(* IEC 61131-3 sources: CNC-Cell-Simulator/source/plc (part 2) *)

PROGRAM CellMain
  VAR_EXTERNAL
    R1_state : INT;
    R1_fault : INT;
    CONV_state : INT;
    CONV_fault : INT;
    R2_state : INT;
    R2_fault : INT;
    SUP_state : INT;
    SAF_state : INT;
    R1_JobNo : INT;
    R1_Start : BOOL;
    R1_Done : BOOL;
    R1_CP_1_Trig : BOOL;
    R1_CP_1_Done : BOOL;
    R1_CP_1_Valid : BOOL;
    R1_CP_1_Cam : BOOL;
    R1_CP_1_Also : BOOL;
    R1_CP_2_Trig : BOOL;
    R1_CP_2_Done : BOOL;
    R1_CP_2_Valid : BOOL;
    R1_CP_2_Cam : BOOL;
    CONV_CP_2_Trig : BOOL;
    CONV_CP_2_Done : BOOL;
    CONV_CP_2_Valid : BOOL;
    CONV_CP_2_Cam : BOOL;
    CONV_CP_3_Trig : BOOL;
    CONV_CP_3_Done : BOOL;
    CONV_CP_3_Valid : BOOL;
    CONV_CP_3_Cam : BOOL;
    R2_JobNo : INT;
    R2_Start : BOOL;
    R2_Done : BOOL;
    R2_CP_4_Trig : BOOL;
    R2_CP_4_Done : BOOL;
    R2_CP_4_Valid : BOOL;
    R2_CP_4_Cam : BOOL;
    R2_CP_5_Trig : BOOL;
    R2_CP_5_Done : BOOL;
    R2_CP_5_Valid : BOOL;
    R2_CP_5_Cam : BOOL;
    R2_CP_3_Trig : BOOL;
    R2_CP_3_Done : BOOL;
    R2_CP_3_Valid : BOOL;
    R2_CP_3_Cam : BOOL;
    HMI_auto : BOOL;
    R1_home : BOOL;
    CNC_ready : BOOL;
    ZS_32_in : BOOL;
    ZS_32 : BOOL;
    SC_01_prot : BOOL;
    GR_21A_in : BOOL;
    GR_21A : BOOL;
    CNC_done : BOOL;
    CNC_empty : BOOL;
    ZS_33_in : BOOL;
    ZS_33 : BOOL;
    ZS_31_in : BOOL;
    ZS_31 : BOOL;
    PS_36_in : BOOL;
    PS_36 : BOOL;
    GR_21B_in : BOOL;
    GR_21B : BOOL;
    ZS_34_in : BOOL;
    ZS_34 : BOOL;
    ZS_35_in : BOOL;
    ZS_35 : BOOL;
    R1_clearCnc : BOOL;
    CNC_run : BOOL;
    ENC_43_in : BOOL;
    ENC_43 : BOOL;
    R1_clearConv : BOOL;
    HMI_loaded : BOOL;
    R2_clearConv : BOOL;
    PE_42_in : BOOL;
    PE_42 : BOOL;
    ROI_C : BOOL;
    R2_home : BOOL;
    GAUGE_zeroed : BOOL;
    GAUGE_due : BOOL;
    GAUGE_due_restart : BOOL;
    GR_51_in : BOOL;
    GR_51 : BOOL;
    R2_clearGauge : BOOL;
    GAUGE_valid : BOOL;
    GAUGE_ok : BOOL;
    SC_02_prot : BOOL;
    CAM_2_slot : BOOL;
    outCount : INT;
    PE_65_in : BOOL;
    PE_65 : BOOL;
    ESTOP : BOOL;
    R1_safeStop : BOOL;
    R2_safeStop : BOOL;
    SC_01_warn : BOOL;
    SC_02_warn : BOOL;
    GAUGE_warn : BOOL;
    PX_11_in : BOOL;
    PX_11 : BOOL;
    PE_41_in : BOOL;
    PE_41 : BOOL;
    PX_52_in : BOOL;
    PX_52 : BOOL;
    PX_64_in : BOOL;
    PX_64 : BOOL;
    HMI_clear : BOOL;
    E_HMI_clear : BOOL;
    HMI_verify : BOOL;
    L_HMI_verify : BOOL;
    VERIFY_pass : BOOL;
    L_VERIFY_pass : BOOL;
    HMI_reset : BOOL;
    L_HMI_reset : BOOL;
    VERIFY_fail : BOOL;
    L_VERIFY_fail : BOOL;
    HMI_safety : BOOL;
    L_HMI_safety : BOOL;
    HMI_release : BOOL;
    L_HMI_release : BOOL;
    HMI_tool : BOOL;
    L_HMI_tool : BOOL;
    HB : BOOL;
    partPlaced : BOOL;
    pickAllowed : BOOL;
    partPicked : BOOL;
    consecNok : INT;
    QH : BOOL;
    toolCount : INT;
    mismatches : INT;
    CAM_FAULT : BOOL;
    COMM_LOST : BOOL;
    mmPending : INT;
    mmClear : BOOL;
    BELT_motor : BOOL;
    LT_53 : BOOL;
    LT_01_red : BOOL;
    LT_01_amber : BOOL;
    LT_01_green : BOOL;
    V_partPlaced : BOOL;
    V_pickAllowed : BOOL;
    V_partPicked : BOOL;
    V_consecNok : INT;
    V_QH : BOOL;
    V_toolCount : INT;
    V_mismatches : INT;
    V_CAM_FAULT : BOOL;
    TR_N : INT;
    TR_00 : INT;
    TR_01 : INT;
    TR_02 : INT;
    TR_03 : INT;
    TR_04 : INT;
    TR_05 : INT;
    TR_06 : INT;
    TR_07 : INT;
    TR_08 : INT;
    TR_09 : INT;
    TR_10 : INT;
    TR_11 : INT;
    TR_12 : INT;
    TR_13 : INT;
    TR_14 : INT;
    TR_15 : INT;
    TR_16 : INT;
    TR_17 : INT;
    TR_18 : INT;
    TR_19 : INT;
    TR_20 : INT;
    TR_21 : INT;
    TR_22 : INT;
    TR_23 : INT;
    TR_24 : INT;
    TR_25 : INT;
    TR_26 : INT;
    TR_27 : INT;
    TR_28 : INT;
    TR_29 : INT;
    TR_30 : INT;
    TR_31 : INT;
  END_VAR
  VAR
    fbR1S2 : FB_R1S2;
    fbCONV : FB_CONV;
    fbR2S2 : FB_R2S2;
    fbSUP : FB_SUP;
    fbSAF : FB_SAF;
    hbT : TON;
    hbLast : BOOL;
    n : INT;
    oldest : INT;
    best : TIME;
    db_ZS_32 : TON;
    db_GR_21A : TON;
    db_ZS_33 : TON;
    db_ZS_31 : TON;
    db_PS_36 : TON;
    db_GR_21B : TON;
    db_ZS_34 : TON;
    db_ZS_35 : TON;
    db_ENC_43 : TON;
    db_PE_42 : TON;
    db_GR_51 : TON;
    db_PX_11 : TON;
    db_PE_41 : TON;
    db_PX_52 : TON;
    db_PX_64 : TON;
    rt_PE_65 : R_TRIG;
    rt_HMI_clear : R_TRIG;
    rt_HMI_verify : R_TRIG;
    rt_VERIFY_pass : R_TRIG;
    rt_HMI_reset : R_TRIG;
    rt_VERIFY_fail : R_TRIG;
    rt_HMI_safety : R_TRIG;
    rt_HMI_release : R_TRIG;
    rt_HMI_tool : R_TRIG;
    mmOn1 : BOOL;
    mmT1 : TON;
    mmOn2 : BOOL;
    mmT2 : TON;
    mmOn3 : BOOL;
    mmT3 : TON;
    tm_GAUGE_due : TON;
    trBuf : ARRAY[0..31] OF INT;
    trI : INT;
    trL_R1 : INT;
    trL_CONV : INT;
    trL_R2 : INT;
    trL_SUP : INT;
    trL_SAF : INT;
  END_VAR
  (* 1. inputs: heartbeat, debounce, latches, mismatch window, PLC timers *)
  hbT(IN := HB = hbLast, PT := T#500ms); hbLast := HB; COMM_LOST := hbT.Q;
  db_ZS_32(IN := ZS_32_in <> ZS_32, PT := T#50ms); IF db_ZS_32.Q THEN ZS_32 := ZS_32_in; END_IF;
  db_GR_21A(IN := GR_21A_in <> GR_21A, PT := T#50ms); IF db_GR_21A.Q THEN GR_21A := GR_21A_in; END_IF;
  db_ZS_33(IN := ZS_33_in <> ZS_33, PT := T#50ms); IF db_ZS_33.Q THEN ZS_33 := ZS_33_in; END_IF;
  db_ZS_31(IN := ZS_31_in <> ZS_31, PT := T#50ms); IF db_ZS_31.Q THEN ZS_31 := ZS_31_in; END_IF;
  db_PS_36(IN := PS_36_in <> PS_36, PT := T#50ms); IF db_PS_36.Q THEN PS_36 := PS_36_in; END_IF;
  db_GR_21B(IN := GR_21B_in <> GR_21B, PT := T#50ms); IF db_GR_21B.Q THEN GR_21B := GR_21B_in; END_IF;
  db_ZS_34(IN := ZS_34_in <> ZS_34, PT := T#50ms); IF db_ZS_34.Q THEN ZS_34 := ZS_34_in; END_IF;
  db_ZS_35(IN := ZS_35_in <> ZS_35, PT := T#50ms); IF db_ZS_35.Q THEN ZS_35 := ZS_35_in; END_IF;
  db_ENC_43(IN := ENC_43_in <> ENC_43, PT := T#50ms); IF db_ENC_43.Q THEN ENC_43 := ENC_43_in; END_IF;
  db_PE_42(IN := PE_42_in <> PE_42, PT := T#50ms); IF db_PE_42.Q THEN PE_42 := PE_42_in; END_IF;
  db_GR_51(IN := GR_51_in <> GR_51, PT := T#50ms); IF db_GR_51.Q THEN GR_51 := GR_51_in; END_IF;
  db_PX_11(IN := PX_11_in <> PX_11, PT := T#50ms); IF db_PX_11.Q THEN PX_11 := PX_11_in; END_IF;
  db_PE_41(IN := PE_41_in <> PE_41, PT := T#50ms); IF db_PE_41.Q THEN PE_41 := PE_41_in; END_IF;
  db_PX_52(IN := PX_52_in <> PX_52, PT := T#50ms); IF db_PX_52.Q THEN PX_52 := PX_52_in; END_IF;
  db_PX_64(IN := PX_64_in <> PX_64, PT := T#50ms); IF db_PX_64.Q THEN PX_64 := PX_64_in; END_IF;
  rt_PE_65(CLK := PE_65_in); IF rt_PE_65.Q THEN PE_65 := TRUE; END_IF;
  rt_HMI_clear(CLK := HMI_clear); E_HMI_clear := rt_HMI_clear.Q;
  rt_HMI_verify(CLK := HMI_verify); IF rt_HMI_verify.Q THEN L_HMI_verify := TRUE; END_IF;
  rt_VERIFY_pass(CLK := VERIFY_pass); IF rt_VERIFY_pass.Q THEN L_VERIFY_pass := TRUE; END_IF;
  rt_HMI_reset(CLK := HMI_reset); IF rt_HMI_reset.Q THEN L_HMI_reset := TRUE; END_IF;
  rt_VERIFY_fail(CLK := VERIFY_fail); IF rt_VERIFY_fail.Q THEN L_VERIFY_fail := TRUE; END_IF;
  rt_HMI_safety(CLK := HMI_safety); IF rt_HMI_safety.Q THEN L_HMI_safety := TRUE; END_IF;
  rt_HMI_release(CLK := HMI_release); IF rt_HMI_release.Q THEN L_HMI_release := TRUE; END_IF;
  rt_HMI_tool(CLK := HMI_tool); IF rt_HMI_tool.Q THEN L_HMI_tool := TRUE; END_IF;
  IF mmClear THEN mmOn1 := FALSE; mmOn2 := FALSE; mmOn3 := FALSE; mmClear := FALSE; END_IF;
  WHILE mmPending > 0 DO (* a new mismatch event: a free place, or the oldest one is replaced *)
    oldest := 0; best := T#0ms;
    IF oldest >= 0 AND NOT mmOn1 THEN oldest := -1; ELSIF oldest >= 0 AND mmT1.ET >= best THEN best := mmT1.ET; oldest := 1; END_IF;
    IF oldest >= 0 AND NOT mmOn2 THEN oldest := -2; ELSIF oldest >= 0 AND mmT2.ET >= best THEN best := mmT2.ET; oldest := 2; END_IF;
    IF oldest >= 0 AND NOT mmOn3 THEN oldest := -3; ELSIF oldest >= 0 AND mmT3.ET >= best THEN best := mmT3.ET; oldest := 3; END_IF;
    IF oldest < 0 THEN oldest := -oldest; END_IF;
    IF oldest = 1 THEN mmOn1 := TRUE; mmT1(IN := FALSE); END_IF;
    IF oldest = 2 THEN mmOn2 := TRUE; mmT2(IN := FALSE); END_IF;
    IF oldest = 3 THEN mmOn3 := TRUE; mmT3(IN := FALSE); END_IF;
    mmPending := mmPending - 1;
  END_WHILE;
  n := 0;
  mmT1(IN := mmOn1, PT := T#600000ms); IF mmT1.Q THEN mmOn1 := FALSE; mmT1(IN := FALSE); END_IF; IF mmOn1 THEN n := n + 1; END_IF;
  mmT2(IN := mmOn2, PT := T#600000ms); IF mmT2.Q THEN mmOn2 := FALSE; mmT2(IN := FALSE); END_IF; IF mmOn2 THEN n := n + 1; END_IF;
  mmT3(IN := mmOn3, PT := T#600000ms); IF mmT3.Q THEN mmOn3 := FALSE; mmT3(IN := FALSE); END_IF; IF mmOn3 THEN n := n + 1; END_IF;
  mismatches := n;
  IF GAUGE_due_restart THEN tm_GAUGE_due(IN := FALSE); GAUGE_due_restart := FALSE; END_IF;
  tm_GAUGE_due(IN := GAUGE_zeroed, PT := T#14400000ms); GAUGE_due := tm_GAUGE_due.Q;

  (* 2. machines in a fixed order; the urgent supervisor first and after every other machine *)
  fbSUP(); IF SUP_state <> trL_SUP THEN trL_SUP := SUP_state; trBuf[trI MOD 32] := 400 + SUP_state; trI := trI + 1; IF trI >= 32000 THEN trI := 0; END_IF; END_IF;
  fbSAF(); IF SAF_state <> trL_SAF THEN trL_SAF := SAF_state; trBuf[trI MOD 32] := 500 + SAF_state; trI := trI + 1; IF trI >= 32000 THEN trI := 0; END_IF; END_IF;
  fbR1S2(); IF R1_state <> trL_R1 THEN trL_R1 := R1_state; trBuf[trI MOD 32] := 100 + R1_state; trI := trI + 1; IF trI >= 32000 THEN trI := 0; END_IF; END_IF;
  fbSUP(); IF SUP_state <> trL_SUP THEN trL_SUP := SUP_state; trBuf[trI MOD 32] := 400 + SUP_state; trI := trI + 1; IF trI >= 32000 THEN trI := 0; END_IF; END_IF;
  fbSAF(); IF SAF_state <> trL_SAF THEN trL_SAF := SAF_state; trBuf[trI MOD 32] := 500 + SAF_state; trI := trI + 1; IF trI >= 32000 THEN trI := 0; END_IF; END_IF;
  fbCONV(); IF CONV_state <> trL_CONV THEN trL_CONV := CONV_state; trBuf[trI MOD 32] := 200 + CONV_state; trI := trI + 1; IF trI >= 32000 THEN trI := 0; END_IF; END_IF;
  fbSUP(); IF SUP_state <> trL_SUP THEN trL_SUP := SUP_state; trBuf[trI MOD 32] := 400 + SUP_state; trI := trI + 1; IF trI >= 32000 THEN trI := 0; END_IF; END_IF;
  fbSAF(); IF SAF_state <> trL_SAF THEN trL_SAF := SAF_state; trBuf[trI MOD 32] := 500 + SAF_state; trI := trI + 1; IF trI >= 32000 THEN trI := 0; END_IF; END_IF;
  fbR2S2(); IF R2_state <> trL_R2 THEN trL_R2 := R2_state; trBuf[trI MOD 32] := 300 + R2_state; trI := trI + 1; IF trI >= 32000 THEN trI := 0; END_IF; END_IF;
  IF (L_HMI_release AND QH) THEN QH := FALSE; consecNok := 0; L_HMI_release := FALSE; END_IF; (* rung: tool and offsets checked -> quality hold released *)
  IF (L_HMI_tool AND (R1_state = 12)) THEN toolCount := 0; L_HMI_tool := FALSE; END_IF; (* rung: tool changed -> tool life counter reset *)
  fbSUP(); IF SUP_state <> trL_SUP THEN trL_SUP := SUP_state; trBuf[trI MOD 32] := 400 + SUP_state; trI := trI + 1; IF trI >= 32000 THEN trI := 0; END_IF; END_IF;
  fbSAF(); IF SAF_state <> trL_SAF THEN trL_SAF := SAF_state; trBuf[trI MOD 32] := 500 + SAF_state; trI := trI + 1; IF trI >= 32000 THEN trI := 0; END_IF; END_IF;

  (* 3. outputs *)
  BELT_motor := (CONV_state = 3) AND NOT COMM_LOST;
  LT_53 := (R2_state = 10);
  LT_01_red := (((SUP_state = 3) OR (SUP_state = 4)) OR ((R1_state = 99) OR (CONV_state = 99) OR (R2_state = 99)) OR ((SAF_state = 4) OR (SAF_state = 5)));
  LT_01_amber := (NOT (((SUP_state = 3) OR (SUP_state = 4))) AND NOT (((R1_state = 99) OR (CONV_state = 99) OR (R2_state = 99))) AND NOT (((SAF_state = 4) OR (SAF_state = 5))) AND ((mismatches > 0) OR QH OR (R1_state = 10) OR (R1_state = 11) OR (R1_state = 12) OR GAUGE_warn OR (SAF_state = 2) OR (SAF_state = 3)));
  LT_01_green := (NOT (((SUP_state = 3) OR (SUP_state = 4))) AND NOT (((R1_state = 99) OR (CONV_state = 99) OR (R2_state = 99))) AND NOT (((SAF_state = 4) OR (SAF_state = 5))) AND NOT (((mismatches > 0) OR QH OR (R1_state = 10) OR (R1_state = 11) OR (R1_state = 12) OR GAUGE_warn OR (SAF_state = 2) OR (SAF_state = 3))));
  V_partPlaced := partPlaced;
  V_pickAllowed := pickAllowed;
  V_partPicked := partPicked;
  V_consecNok := consecNok;
  V_QH := QH;
  V_toolCount := toolCount;
  V_mismatches := mismatches;
  V_CAM_FAULT := CAM_FAULT;
  TR_00 := trBuf[0];
  TR_01 := trBuf[1];
  TR_02 := trBuf[2];
  TR_03 := trBuf[3];
  TR_04 := trBuf[4];
  TR_05 := trBuf[5];
  TR_06 := trBuf[6];
  TR_07 := trBuf[7];
  TR_08 := trBuf[8];
  TR_09 := trBuf[9];
  TR_10 := trBuf[10];
  TR_11 := trBuf[11];
  TR_12 := trBuf[12];
  TR_13 := trBuf[13];
  TR_14 := trBuf[14];
  TR_15 := trBuf[15];
  TR_16 := trBuf[16];
  TR_17 := trBuf[17];
  TR_18 := trBuf[18];
  TR_19 := trBuf[19];
  TR_20 := trBuf[20];
  TR_21 := trBuf[21];
  TR_22 := trBuf[22];
  TR_23 := trBuf[23];
  TR_24 := trBuf[24];
  TR_25 := trBuf[25];
  TR_26 := trBuf[26];
  TR_27 := trBuf[27];
  TR_28 := trBuf[28];
  TR_29 := trBuf[29];
  TR_30 := trBuf[30];
  TR_31 := trBuf[31];
  TR_N := trI;
END_PROGRAM

CONFIGURATION Config0
  VAR_GLOBAL (* inputs from the plant (Modbus bridge, A3.3) *)
    R1_Done AT %IX100.0 : BOOL; (* job done, held until Start is low *)
    R1_CP_1_Done AT %IX100.1 : BOOL; (* camera answer for CP-1 ready, held until Trig is low *)
    R1_CP_1_Valid AT %IX100.2 : BOOL; (* CAM-1 image valid *)
    R1_CP_1_Cam AT %IX100.3 : BOOL; (* CAM-1 / ROI-A: Input pallet present and seated *)
    R1_CP_1_Also AT %IX100.4 : BOOL; (* CAM-1: CAM-1.part *)
    R1_CP_2_Done AT %IX100.5 : BOOL; (* camera answer for CP-2 ready, held until Trig is low *)
    R1_CP_2_Valid AT %IX100.6 : BOOL; (* CAM-1 image valid *)
    R1_CP_2_Cam AT %IX100.7 : BOOL; (* CAM-1 / ROI-B: Part at conveyor entry *)
    CONV_CP_2_Done AT %IX101.0 : BOOL; (* camera answer for CP-2 ready, held until Trig is low *)
    CONV_CP_2_Valid AT %IX101.1 : BOOL; (* CAM-1 image valid *)
    CONV_CP_2_Cam AT %IX101.2 : BOOL; (* CAM-1 / ROI-B: Part at conveyor entry *)
    CONV_CP_3_Done AT %IX101.3 : BOOL; (* camera answer for CP-3 ready, held until Trig is low *)
    CONV_CP_3_Valid AT %IX101.4 : BOOL; (* CAM-2 image valid *)
    CONV_CP_3_Cam AT %IX101.5 : BOOL; (* CAM-2 / ROI-C: Part at the end stop *)
    R2_Done AT %IX101.6 : BOOL; (* job done, held until Start is low *)
    R2_CP_4_Done AT %IX101.7 : BOOL; (* camera answer for CP-4 ready, held until Trig is low *)
    R2_CP_4_Valid AT %IX102.0 : BOOL; (* CAM-2 image valid *)
    R2_CP_4_Cam AT %IX102.1 : BOOL; (* CAM-2 / ROI-D: Output pallet present *)
    R2_CP_5_Done AT %IX102.2 : BOOL; (* camera answer for CP-5 ready, held until Trig is low *)
    R2_CP_5_Valid AT %IX102.3 : BOOL; (* CAM-2 image valid *)
    R2_CP_5_Cam AT %IX102.4 : BOOL; (* CAM-2 / ROI-E: Part in gauge nest *)
    R2_CP_3_Done AT %IX102.5 : BOOL; (* camera answer for CP-3 ready, held until Trig is low *)
    R2_CP_3_Valid AT %IX102.6 : BOOL; (* CAM-2 image valid *)
    R2_CP_3_Cam AT %IX102.7 : BOOL; (* CAM-2 / ROI-C: Part at the end stop *)
    HMI_auto AT %IX103.0 : BOOL; (* HMI.auto *)
    R1_home AT %IX103.1 : BOOL; (* R1.home *)
    CNC_ready AT %IX103.2 : BOOL; (* CNC.ready *)
    ZS_32_in AT %IX103.3 : BOOL; (* ZS-32, raw *)
    SC_01_prot AT %IX103.4 : BOOL; (* SC-01.prot *)
    GR_21A_in AT %IX103.5 : BOOL; (* GR-21A, raw *)
    CNC_done AT %IX103.6 : BOOL; (* CNC.done *)
    CNC_empty AT %IX103.7 : BOOL; (* CNC.empty *)
    ZS_33_in AT %IX104.0 : BOOL; (* ZS-33, raw *)
    ZS_31_in AT %IX104.1 : BOOL; (* ZS-31, raw *)
    PS_36_in AT %IX104.2 : BOOL; (* PS-36, raw *)
    GR_21B_in AT %IX104.3 : BOOL; (* GR-21B, raw *)
    ZS_34_in AT %IX104.4 : BOOL; (* ZS-34, raw *)
    ZS_35_in AT %IX104.5 : BOOL; (* ZS-35, raw *)
    R1_clearCnc AT %IX104.6 : BOOL; (* R1.clearCnc *)
    CNC_run AT %IX104.7 : BOOL; (* CNC.run *)
    ENC_43_in AT %IX105.0 : BOOL; (* ENC-43, raw *)
    R1_clearConv AT %IX105.1 : BOOL; (* R1.clearConv *)
    HMI_loaded AT %IX105.2 : BOOL; (* HMI.loaded *)
    R2_clearConv AT %IX105.3 : BOOL; (* R2.clearConv *)
    PE_42_in AT %IX105.4 : BOOL; (* PE-42, raw *)
    ROI_C AT %IX105.5 : BOOL; (* ROI-C *)
    R2_home AT %IX105.6 : BOOL; (* R2.home *)
    GAUGE_zeroed AT %IX105.7 : BOOL; (* GAUGE.zeroed *)
    GR_51_in AT %IX106.0 : BOOL; (* GR-51, raw *)
    R2_clearGauge AT %IX106.1 : BOOL; (* R2.clearGauge *)
    GAUGE_valid AT %IX106.2 : BOOL; (* GAUGE.valid *)
    GAUGE_ok AT %IX106.3 : BOOL; (* GAUGE.ok *)
    SC_02_prot AT %IX106.4 : BOOL; (* SC-02.prot *)
    CAM_2_slot AT %IX106.5 : BOOL; (* CAM-2.slot *)
    outCount AT %IW100 : INT; (* outCount *)
    PE_65_in AT %IX106.6 : BOOL; (* PE-65, raw *)
    ESTOP AT %IX106.7 : BOOL; (* ESTOP *)
    R1_safeStop AT %IX107.0 : BOOL; (* R1.safeStop *)
    R2_safeStop AT %IX107.1 : BOOL; (* R2.safeStop *)
    SC_01_warn AT %IX107.2 : BOOL; (* SC-01.warn *)
    SC_02_warn AT %IX107.3 : BOOL; (* SC-02.warn *)
    GAUGE_warn AT %IX107.4 : BOOL; (* GAUGE.warn *)
    PX_11_in AT %IX107.5 : BOOL; (* PX-11, raw *)
    PE_41_in AT %IX107.6 : BOOL; (* PE-41, raw *)
    PX_52_in AT %IX107.7 : BOOL; (* PX-52, raw *)
    PX_64_in AT %IX108.0 : BOOL; (* PX-64, raw *)
    HMI_clear AT %IX108.1 : BOOL; (* HMI.clear (button) *)
    HMI_verify AT %IX108.2 : BOOL; (* HMI.verify (button) *)
    VERIFY_pass AT %IX108.3 : BOOL; (* VERIFY.pass (button) *)
    HMI_reset AT %IX108.4 : BOOL; (* HMI.reset (button) *)
    VERIFY_fail AT %IX108.5 : BOOL; (* VERIFY.fail (button) *)
    HMI_safety AT %IX108.6 : BOOL; (* HMI.safety (button) *)
    HMI_release AT %IX108.7 : BOOL; (* HMI.release (button) *)
    HMI_tool AT %IX109.0 : BOOL; (* HMI.tool (button) *)
    HB AT %IX109.1 : BOOL; (* heartbeat, toggled by the bridge *)
  END_VAR
  VAR_GLOBAL (* outputs to the plant *)
    R1_state AT %QW100 : INT; (* state of R1 (codes in FB_R1S2) *)
    R1_fault AT %QW101 : INT; (* fault code of R1, 0 = none *)
    CONV_state AT %QW102 : INT; (* state of CONV (codes in FB_CONV) *)
    CONV_fault AT %QW103 : INT; (* fault code of CONV, 0 = none *)
    R2_state AT %QW104 : INT; (* state of R2 (codes in FB_R2S2) *)
    R2_fault AT %QW105 : INT; (* fault code of R2, 0 = none *)
    SUP_state AT %QW106 : INT; (* state of SUP (codes in FB_SUP) *)
    SAF_state AT %QW107 : INT; (* state of SAF (codes in FB_SAF) *)
    R1_JobNo AT %QW108 : INT; (* job number (order of M.JOBS, from 1; 0 = no job) *)
    R1_Start AT %QX100.0 : BOOL; (* job start (handshake: Start, Done, Start low, Done low) *)
    R1_CP_1_Trig AT %QX100.1 : BOOL; (* camera trigger for CP-1 *)
    R1_CP_2_Trig AT %QX100.2 : BOOL; (* camera trigger for CP-2 *)
    CONV_CP_2_Trig AT %QX100.3 : BOOL; (* camera trigger for CP-2 *)
    CONV_CP_3_Trig AT %QX100.4 : BOOL; (* camera trigger for CP-3 *)
    R2_JobNo AT %QW109 : INT; (* job number (order of M.JOBS, from 1; 0 = no job) *)
    R2_Start AT %QX100.5 : BOOL; (* job start (handshake: Start, Done, Start low, Done low) *)
    R2_CP_4_Trig AT %QX100.6 : BOOL; (* camera trigger for CP-4 *)
    R2_CP_5_Trig AT %QX100.7 : BOOL; (* camera trigger for CP-5 *)
    R2_CP_3_Trig AT %QX101.0 : BOOL; (* camera trigger for CP-3 *)
    BELT_motor AT %QX101.1 : BOOL; (* conveyor motor ON *)
    LT_53 AT %QX101.2 : BOOL; (* blue beacon: output pallet ready for pickup *)
    LT_01_red AT %QX101.3 : BOOL; (* stack light red *)
    LT_01_amber AT %QX101.4 : BOOL; (* stack light amber *)
    LT_01_green AT %QX101.5 : BOOL; (* stack light green *)
    V_partPlaced AT %QX101.6 : BOOL; (* copy of partPlaced *)
    V_pickAllowed AT %QX101.7 : BOOL; (* copy of pickAllowed *)
    V_partPicked AT %QX102.0 : BOOL; (* copy of partPicked *)
    V_consecNok AT %QW110 : INT; (* copy of consecNok *)
    V_QH AT %QX102.1 : BOOL; (* copy of QH *)
    V_toolCount AT %QW111 : INT; (* copy of toolCount *)
    V_mismatches AT %QW112 : INT; (* copy of mismatches *)
    V_CAM_FAULT AT %QX102.2 : BOOL; (* copy of CAM_FAULT *)
    TR_N AT %QW113 : INT; (* state changes so far, modulo 32000 *)
    TR_00 AT %QW114 : INT; (* state change ring: machine number x 100 + state code *)
    TR_01 AT %QW115 : INT;
    TR_02 AT %QW116 : INT;
    TR_03 AT %QW117 : INT;
    TR_04 AT %QW118 : INT;
    TR_05 AT %QW119 : INT;
    TR_06 AT %QW120 : INT;
    TR_07 AT %QW121 : INT;
    TR_08 AT %QW122 : INT;
    TR_09 AT %QW123 : INT;
    TR_10 AT %QW124 : INT;
    TR_11 AT %QW125 : INT;
    TR_12 AT %QW126 : INT;
    TR_13 AT %QW127 : INT;
    TR_14 AT %QW128 : INT;
    TR_15 AT %QW129 : INT;
    TR_16 AT %QW130 : INT;
    TR_17 AT %QW131 : INT;
    TR_18 AT %QW132 : INT;
    TR_19 AT %QW133 : INT;
    TR_20 AT %QW134 : INT;
    TR_21 AT %QW135 : INT;
    TR_22 AT %QW136 : INT;
    TR_23 AT %QW137 : INT;
    TR_24 AT %QW138 : INT;
    TR_25 AT %QW139 : INT;
    TR_26 AT %QW140 : INT;
    TR_27 AT %QW141 : INT;
    TR_28 AT %QW142 : INT;
    TR_29 AT %QW143 : INT;
    TR_30 AT %QW144 : INT;
    TR_31 AT %QW145 : INT;
  END_VAR
  VAR_GLOBAL (* internal *)
    ZS_32 : BOOL; (* ZS-32, debounced *)
    GR_21A : BOOL; (* GR-21A, debounced *)
    ZS_33 : BOOL; (* ZS-33, debounced *)
    ZS_31 : BOOL; (* ZS-31, debounced *)
    PS_36 : BOOL; (* PS-36, debounced *)
    GR_21B : BOOL; (* GR-21B, debounced *)
    ZS_34 : BOOL; (* ZS-34, debounced *)
    ZS_35 : BOOL; (* ZS-35, debounced *)
    ENC_43 : BOOL; (* ENC-43, debounced *)
    PE_42 : BOOL; (* PE-42, debounced *)
    GAUGE_due : BOOL; (* PLC timer (M.PLC.timers) *)
    GAUGE_due_restart : BOOL; (* restart GAUGE.due *)
    GR_51 : BOOL; (* GR-51, debounced *)
    PE_65 : BOOL; (* PE-65, latched on the rising edge *)
    PX_11 : BOOL; (* PX-11, debounced *)
    PE_41 : BOOL; (* PE-41, debounced *)
    PX_52 : BOOL; (* PX-52, debounced *)
    PX_64 : BOOL; (* PX-64, debounced *)
    E_HMI_clear : BOOL; (* rising edge of HMI.clear in this scan *)
    L_HMI_verify : BOOL; (* HMI.verify, latched until a transition reads it *)
    L_VERIFY_pass : BOOL; (* VERIFY.pass, latched until a transition reads it *)
    L_HMI_reset : BOOL; (* HMI.reset, latched until a transition reads it *)
    L_VERIFY_fail : BOOL; (* VERIFY.fail, latched until a transition reads it *)
    L_HMI_safety : BOOL; (* HMI.safety, latched until a transition reads it *)
    L_HMI_release : BOOL; (* HMI.release, latched until a transition reads it *)
    L_HMI_tool : BOOL; (* HMI.tool, latched until a transition reads it *)
    partPlaced : BOOL; (* partPlaced *)
    pickAllowed : BOOL; (* pickAllowed *)
    partPicked : BOOL; (* partPicked *)
    mismatches : INT; (* mismatches *)
    CAM_FAULT : BOOL; (* CAM_FAULT *)
    COMM_LOST : BOOL; (* no heartbeat for M.PLC.heartbeatTimeout *)
    mmPending : INT; (* mismatch events to add to the window *)
    mmClear : BOOL; (* clear the mismatch window *)
  END_VAR
  VAR_GLOBAL RETAIN (* kept over a cold restart (M.PLC.retain) *)
    consecNok : INT; (* consecNok *)
    QH : BOOL; (* QH *)
    toolCount : INT; (* toolCount *)
  END_VAR
  RESOURCE Res0 ON PLC
    TASK MainTask (INTERVAL := T#10ms, PRIORITY := 0);
    PROGRAM Main WITH MainTask : CellMain;
  END_RESOURCE
END_CONFIGURATION
